FUNCTION_BLOCK tonnnnblock
VAR_INPUT
	in:BOOL;
	pt:TIME;
	
END_VAR
VAR_OUTPUT
	out:BOOL;
	et:TIME;
	
END_VAR
VAR
	tstarttime:TIME;
	brunning:BOOL;
END_VAR

IF in THEN
	IF NOT brunning THEN
		tstarttime :=TIME();
		brunning :=TRUE;
		et :=T#0MS;
		out :=FALSE;
	ELSE
		ET := TIME()-tstarttime;
		IF et>=pt THEN
			et:=pt;
			out:=TRUE;
			
		END_IF
	END_IF
ELSE
	brunning :=FALSE;
	et:= T#0MS;
	out:=FALSE;
END_IF

END_FUNCTION_BLOCK

(* stored: Version 1.1.0.1, ProductVersion 3.1.4024.16
   POU tonnnnblock: Id {6a0c1958-6b51-4ffc-a521-727268d0e81c}, SpecialFunc None *)
